Fanuc KAREL source: ks00047.KL

-- PROVISIONAL review KL for V770-1; original PC SHA256 066faac0632960a6b78cb33639a72b34572fce25cad80f0cfe03e270c7699108
-- Incomplete behavior may be omitted. Consult companion uncertainty JSON. Do not deploy.
PROGRAM KS00047
%NOLOCKGROUP
BEGIN
  -- UNRESOLVED_PC offsets 5-13; opcodes 3F,75
  -- UNRESOLVED_PC offsets 18-27; opcodes 3F,75
  -- UNRESOLVED_PC offsets 32-45; opcodes 22,1D,23
  -- UNRESOLVED_PC offsets 50-54; opcodes 7F
END KS00047
